// TIA Portal project "Project1" (V20)

(* hardware
DEVICE "S7-1500/ET200MP station_1"  S7-1500 station
   slot 0: "Rail_0"  Rack  6ES7 590-1***0-0AA0
   slot 1: "PLC_2"  CPU 1515F-2 PN  6ES7 515-2FM01-0AB0  V2.9
      slot 3: "CPU display_1"  6ES7591-1BA00-0AA0
      slot 32768: "PROFINET interface_1"  X1
         slot 32769: "Port_1"  X1 P1
         slot 32770: "Port_2"  X1 P2
      slot 33024: "PROFINET interface_2"  X2
         slot 33025: "Port_1"  X2 P1
      slot 34817: "Virtual CP interface port_1"  Virtual CP interface port  Virtual CP interface port
   slot 2: "DI 16x24VDC BA_1"  DI 16x24VDC BA  6ES7 521-1BH10-0AA0  V1.1
   slot 3: "DQ 16x24VDC/0.5A BA_1"  DQ 16x24VDC/0.5A BA  6ES7 522-1BH10-0AA0  V1.1
DEVICE "HMI_1"  KTP700 Basic PN
   slot 0: "HMI_1"  KTP700 Basic PN  6AV2 123-2GB03-0AX0  17.0.0.0
   slot 1: "HMI_RT_1"  KTP700 Basic PN  6AV2 123-2GB03-0AX0  17.0.0.0
   slot 5: "HMI_1.IE_CP_1"  PROFINET Interface  17.0.0.0
      slot 1: "PROFINET Interface_1"  PROFINET Interface
         slot 1: "Port_1"  Port
*)

// ===== PLC "PLC_2"  CPU 1515F-2 PN =====

VAR_GLOBAL   // PLC tag table "Default tag table"
   "KM_Moteur" AT %Q0.0 : Bool;
   "BP_Marche" AT %M0.0 : Bool;
   "BP_Arret_OK" AT %M0.1 : Bool;
   "Niveau_Cuve" AT %MD20 : Real;
   "Vitesse_Pompe" AT %MD24 : Real;
   "Vanne_Vidange" AT %M0.3 : Bool;
   "Cuve_Pleine" AT %M0.2 : Bool;
   "Demande_Production" AT %MD28 : Real;
   "Debit_Sortie" AT %MD32 : Real;
   "Delta_Niveau_Sortie" AT %MD36 : Real;
   "Niveau_Cuve_Calcule" AT %MD40 : Real;
   "Demande_Production_Limitee" AT %MD44 : Real;
   "Debit_Entree" AT %MD48 : Real;
   "Delta_Niveau_Entree" AT %MD52 : Real;
   "Debit_Vidange" AT %MD56 : Real;
   "Autorisation_Vidange" AT %M0.4 : Bool;
   "Debit_Sortie_Total" AT %MD60 : Real;
   "Niveau_Apres_Entree" AT %MD64 : Real;
   "Debit_Entree_Theorique" AT %MD68 : Real;
   "Vitesse_Pompe_Manuelle" AT %MD72 : Real;
END_VAR

DATA_BLOCK "Main_Safety_RTG1_DB"   // DB1, F_DB
{ S7_Optimized_Access := 'TRUE' }
NAME : FUSI
VERSION : 0.1
// stored: InstanceOfName Main_Safety_RTG1
"Main_Safety_RTG1"
BEGIN
END_DATA_BLOCK

DATA_BLOCK "FB_Regulation_Niveau_DB"   // DB3
{ S7_Optimized_Access := 'TRUE' }
VERSION : 0.1
// stored: InstanceOfName FB_Regulation_Niveau
"FB_Regulation_Niveau"
BEGIN
END_DATA_BLOCK

FUNCTION_BLOCK "Main_Safety_RTG1"   // FB1, F_FBD
{ S7_Optimized_Access := 'TRUE' }
BEGIN
END_FUNCTION_BLOCK

FUNCTION_BLOCK "FB_Regulation_Niveau"   // FB2, LAD
{ S7_Optimized_Access := 'TRUE' }
VERSION : 0.1
   VAR
      Consigne_Niveau : Real := 70.0;
      Mode_Auto : Bool;
      Vitesse_PID : Real;
      PID_Actif : Bool;
      Mode_Manuel : Bool;
      Mode_PID : Int := 3;
      Etat_PID : Int;
   END_VAR
BEGIN

REGION Network 1
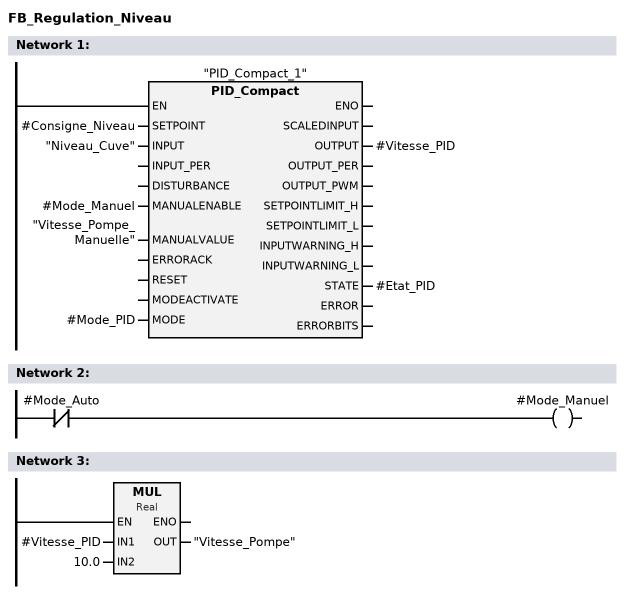
   "PID_Compact_1"(Setpoint := #Consigne_Niveau,   // PID_Compact
                   Input := "Niveau_Cuve",
                   ManualEnable := #Mode_Manuel,
                   ManualValue := "Vitesse_Pompe_Manuelle",
                   Mode := #Mode_PID,
                   Output => #Vitesse_PID,
                   State => #Etat_PID);
END_REGION

REGION Network 2
   RUNG wire#powerrail
      I_Contact( #Mode_Auto )
      Coil( #Mode_Manuel )
   END_RUNG
   // the same network as SCL:
   #Mode_Manuel := NOT #Mode_Auto;
END_REGION

REGION Network 3
   RUNG wire#powerrail
      { S7_Templates := "SrcType := Real" } Mul(in1 := #Vitesse_PID, in2 := 10.0, out => "Vitesse_Pompe")
   END_RUNG
   // the same network as SCL:
   "Vitesse_Pompe" := #Vitesse_PID * 10.0;
END_REGION
END_FUNCTION_BLOCK

ORGANIZATION_BLOCK "Main"   // OB1, LAD, ProgramCycle
TITLE = "Main Program Sweep (Cycle)"
{ S7_Optimized_Access := 'TRUE' }
VERSION : 0.1
   VAR_INPUT
      Initial_Call : Bool;   // Initial call of this OB
      Remanence : Bool;   // =True, if remanent data are available
   END_VAR
BEGIN

REGION Network 1
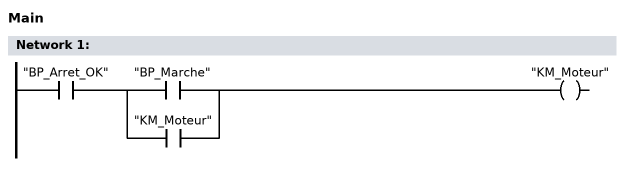
   RUNG wire#powerrail
      Contact( "BP_Arret_OK" )
      wire#w1
      Contact( "BP_Marche" )
      wire#w2
      Coil( "KM_Moteur" )
   END_RUNG
   RUNG wire#w1
      Contact( "KM_Moteur" )
   END_RUNG wire#w2
   // the same network as SCL:
   "KM_Moteur" := "BP_Arret_OK" AND ("BP_Marche" OR "KM_Moteur");
END_REGION
END_ORGANIZATION_BLOCK

ORGANIZATION_BLOCK "OB30_Simulation_Cuve"   // OB30, LAD, CyclicInterrupt
{ S7_Optimized_Access := 'TRUE' }
VERSION : 0.1
   VAR_INPUT
      Initial_Call : Bool;   // Initial call of this OB
      Event_Count : Int;   // Events discarded
   END_VAR
BEGIN

REGION Network 1
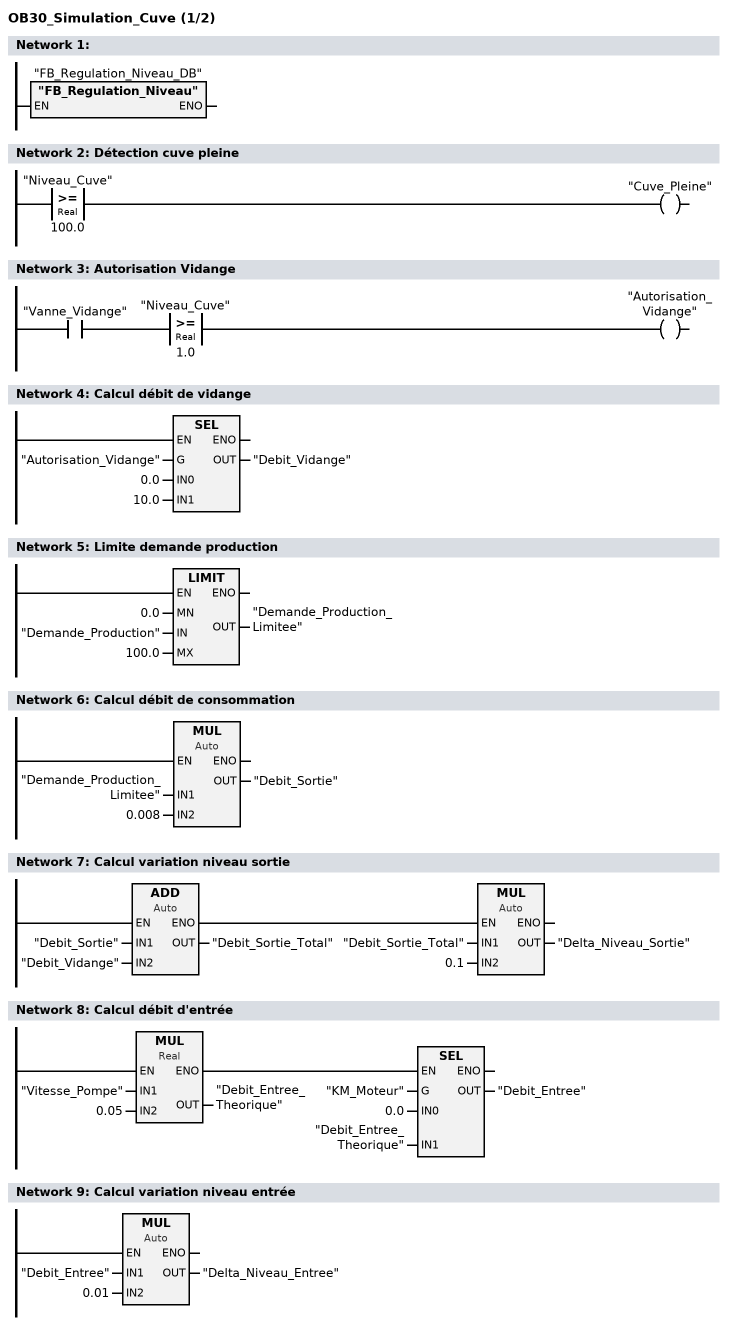
   RUNG wire#powerrail
      "FB_Regulation_Niveau_DB"()
   END_RUNG
   // the same network as SCL:
   "FB_Regulation_Niveau_DB"();   // "FB_Regulation_Niveau"
END_REGION

REGION Network 2: Détection cuve pleine
   RUNG wire#powerrail
      { S7_Templates := "SrcType := Real" } GE_Contact(in1 := "Niveau_Cuve", in2 := 100.0)
      Coil( "Cuve_Pleine" )
   END_RUNG
   // the same network as SCL:
   "Cuve_Pleine" := "Niveau_Cuve" >= 100.0;
END_REGION

REGION Network 3: Autorisation Vidange
   RUNG wire#powerrail
      Contact( "Vanne_Vidange" )
      { S7_Templates := "SrcType := Real" } GE_Contact(in1 := "Niveau_Cuve", in2 := 1.0)
      Coil( "Autorisation_Vidange" )
   END_RUNG
   // the same network as SCL:
   "Autorisation_Vidange" := "Vanne_Vidange" AND ("Niveau_Cuve" >= 1.0);
END_REGION

REGION Network 4: Calcul débit de vidange
   "Debit_Vidange" := SEL(G := "Autorisation_Vidange", IN0 := 0.0, IN1 := 10.0);
END_REGION

REGION Network 5: Limite demande production
   "Demande_Production_Limitee" := LIMIT(MN := 0.0, IN := "Demande_Production", MX := 100.0);
END_REGION

REGION Network 6: Calcul débit de consommation
   RUNG wire#powerrail
      Mul(in1 := "Demande_Production_Limitee", in2 := 0.008, out => "Debit_Sortie")
   END_RUNG
   // the same network as SCL:
   "Debit_Sortie" := "Demande_Production_Limitee" * 0.008;
END_REGION

REGION Network 7: Calcul variation niveau sortie
   RUNG wire#powerrail
      Add(in1 := "Debit_Sortie", in2 := "Debit_Vidange", out => "Debit_Sortie_Total")
      Mul(in1 := "Debit_Sortie_Total", in2 := 0.1, out => "Delta_Niveau_Sortie")
   END_RUNG
   // the same network as SCL:
   "Debit_Sortie_Total" := "Debit_Sortie" + "Debit_Vidange";
   "Delta_Niveau_Sortie" := "Debit_Sortie_Total" * 0.1;
END_REGION

REGION Network 8: Calcul débit d'entrée
   "Debit_Entree_Theorique" := "Vitesse_Pompe" * 0.05;
   "Debit_Entree" := SEL(G := "KM_Moteur", IN0 := 0.0, IN1 := "Debit_Entree_Theorique");
END_REGION

REGION Network 9: Calcul variation niveau entrée
   RUNG wire#powerrail
      Mul(in1 := "Debit_Entree", in2 := 0.01, out => "Delta_Niveau_Entree")
   END_RUNG
   // the same network as SCL:
   "Delta_Niveau_Entree" := "Debit_Entree" * 0.01;
END_REGION

REGION Network 10: Calcul niveau après remplissage
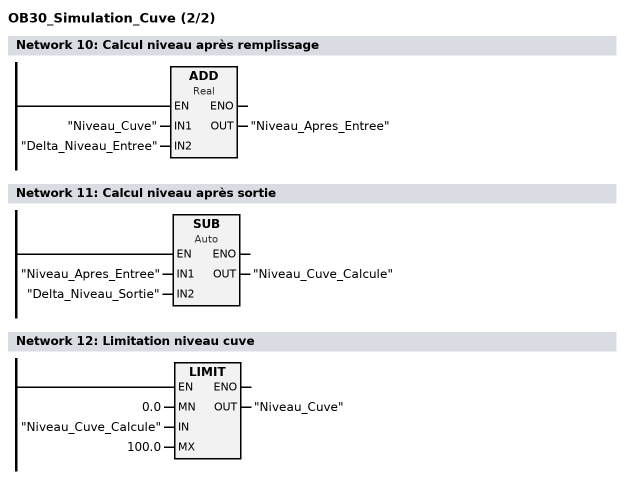
   RUNG wire#powerrail
      { S7_Templates := "SrcType := Real" } Add(in1 := "Niveau_Cuve", in2 := "Delta_Niveau_Entree", out => "Niveau_Apres_Entree")
   END_RUNG
   // the same network as SCL:
   "Niveau_Apres_Entree" := "Niveau_Cuve" + "Delta_Niveau_Entree";
END_REGION

REGION Network 11: Calcul niveau après sortie
   RUNG wire#powerrail
      Sub(in1 := "Niveau_Apres_Entree", in2 := "Delta_Niveau_Sortie", out => "Niveau_Cuve_Calcule")
   END_RUNG
   // the same network as SCL:
   "Niveau_Cuve_Calcule" := "Niveau_Apres_Entree" - "Delta_Niveau_Sortie";
END_REGION

REGION Network 12: Limitation niveau cuve
   "Niveau_Cuve" := LIMIT(MN := 0.0, IN := "Niveau_Cuve_Calcule", MX := 100.0);
END_REGION
END_ORGANIZATION_BLOCK

(* ===== HMI "HMI_RT_1" =====
system functions are stored by id; their names below are inferred from use
connection "HMI_Connection_2": ETHERNET, SMART_S7_1500_OMS
connection "HMI_Connection_3": ETHERNET, SMART_S7_1500_OMS

HMI tags "Default tag table"
   "Vanne_Vidange_HMI" : Bool = PLC Vanne_Vidange AT %M0.3, 1 s
   "BP_Marche" : Bool = PLC BP_Marche AT %M0.0, 1 s
   "BP_Arret_OK" : Bool = PLC BP_Arret_OK AT %M0.1, 1 s
   "KM_Moteur" : Bool = PLC KM_Moteur AT %Q0.0, 1 s
   "Demande_Production_HMI" : Real = PLC Demande_Production AT %MD28, 1 s
   "Niveau_Cuve_HMI" : Real = PLC Niveau_Cuve AT %MD20, 1 s
   "Vitesse_Pompe_Manuelle_HMI" : Real = PLC Vitesse_Pompe_Manuelle AT %MD72, 1 s
   "Mode_Auto_HMI" : Bool = PLC FB_Regulation_Niveau_DB.Mode_Auto AT %DB1.DBX0.0, 1 s
   "Consigne_Niveau_HMI" : Real = PLC FB_Regulation_Niveau_DB.Consigne_Niveau AT %DB1.DBX0.0, 1 s
   "PID_Compact_1_CtrlParamsBackUp_Gain" : Real = PLC PID_Compact_1.CtrlParamsBackUp.Gain, 1 s
   "PID_Compact_1_CtrlParamsBackUp_Ti" : Real = PLC PID_Compact_1.CtrlParamsBackUp.Ti, 1 s
   "PID_Compact_1_Retain_CtrlParams_Gain" : Real = PLC PID_Compact_1.Retain.CtrlParams.Gain, 1 s
   "PID_Compact_1_Retain_CtrlParams_Ti" : Real = PLC PID_Compact_1.Retain.CtrlParams.Ti, 1 s

Template "Template_1" 800x480
   Button "Exit" at 714,429 size 71x50; TextOff 'Exit'; PictureOff "ExitRuntime_KTP700_Basic_DP_TR"; PictureOn "ExitRuntime_KTP700_Basic_DP_TR"
      on Release: StopRuntime(0)
   Button "Template_Button" at 614,429 size 71x50; TextOff 'Text'
   Button "Template_Button_1" at 514,429 size 71x50; TextOff 'Text'
   Button "Template_Button_2" at 414,429 size 71x50; TextOff 'Text'
   Button "Template_Button_3" at 314,429 size 71x50; TextOff 'Text'
   Button "Template_Button_4" at 214,429 size 71x50; TextOff 'Text'
   Button "Alarms" at 114,429 size 71x50; TextOff 'Alarms'; PictureOff "AlarmDisplay_KTP700_Basic_DP_TR"; PictureOn "AlarmDisplay_KTP700_Basic_DP_TR"
      on Release: function_ef3f5d25("Alarm window_Unacknowledged", -1)
   Button "Start screen" at 14,429 size 71x50; TextOff 'Start screen'; PictureOff "NavigateHome_KTP700_Basic_DP_TR"; PictureOn "NavigateHome_KTP700_Basic_DP_TR"
      on Release: ActivateScreen("Root screen", 0)
   SymbolicIOField "Symbolic_IO_Field_Screen" at 93,9 size 600x33; TextOff '0'; TextOn '1'; TextList "TextList_ScreenNames"
      ProcessValue <- "Vanne_Vidange_HMI"
   DateTimeField "HmiScreenItemData" at 695,25 size 105x25
   DateTimeField "HmiScreenItemData_1" at 695,0 size 105x25
   GraphicView "Logo" at 0,0 size 91x51; Picture "Logo of HMI_1"

screen "Root screen" 800x480, template "Template_1"
   on GenerateScreen: SetTag("Vanne_Vidange_HMI", 1)
   TextField "HmiScreenItemData" at 80,225 size 640x25; Text 'Welcome to HMI_1 (KTP700 Basic+ DP)!'

screen "Screen_1" 800x480
   Bar "Bar_1" at 536,85 size 41x217; MinimumValue 0; MaximumValue 100
      ProcessValue <- "Niveau_Cuve_HMI"
   IOField "I/O field_1" at 659,147 size 49x38; FormatPattern 999
      ProcessValue <- "Demande_Production_HMI"
   IOField "I/O field_4" at 85,253 size 96x32; FormatPattern s999999999.999
      ProcessValue <- "Consigne_Niveau_HMI"
   IOField "I/O field_3" at 126,163 size 68x28; FormatPattern s999999999.999
      ProcessValue <- "Vitesse_Pompe_Manuelle_HMI"
   IOField "I/O field_2" at 393,152 size 96x32; FormatPattern s999999999.999
      ProcessValue <- "Niveau_Cuve_HMI"
   Switch "Switch_1" at 126,127 size 57x26; CaptionText 'Switch'; TextOff 'OFF'; TextOn 'ON'
      ProcessValue <- "Mode_Auto_HMI"
   TextField "Text field_2" at 12,127 size 110x20; Text 'AUTO [ON/OFF] :'
   TextField "Text field_3" at 9,163 size 113x20; Text 'MANUAL VALUE :'
   TextField "Text field_4" at 12,253 size 73x20; Text 'SETPOINT :'
   IOField "I/O field_5" at 85,285 size 96x32; FormatPattern s999999999.999
      ProcessValue <- "PID_Compact_1_Retain_CtrlParams_Gain"
   TextField "Text field_5" at 33,291 size 41x20; Text 'Gain :'
   TextField "Text field_6" at 48,317 size 28x20; Text 'Ti :'
   IOField "I/O field_6" at 85,317 size 96x32; FormatPattern s999999999.999
      ProcessValue <- "PID_Compact_1_Retain_CtrlParams_Ti"
   TextField "Text field_7" at 612,93 size 148x23; Text 'WATER DEMAND'
   TextField "Text field_1" at 602,195 size 158x59; Text '0 % No consumption 25 % Low consumption 50 % Medium consumption 75 % High consumption 100 % Maximum consumption'
   TextField "Text field_8" at 39,19 size 164x28; Text 'PUMP SETTINGS'
   TextField "Text field_9" at 55,205 size 128x22; Text 'PI PARAMETERS'
   TextField "Text field_10" at 48,71 size 145x22; Text 'OPERATING MODE'
   Button "Button_1" at 12,436 size 96x32; TextOff 'RUN'
      on Press: SetBit("BP_Marche")
      on Release: ResetBit("BP_Marche")
   Button "Button_2" at 129,437 size 96x32; TextOff 'STOP'
      on Press: ResetBit("BP_Arret_OK")
      on Release: SetBit("BP_Arret_OK")
   Circle "Circle_1" at 76,363 size 67x67
      Appearance <- "KM_Moteur"
   TextField "Text field_11" at 379,399 size 144x23; Text 'DRAIN CONTROL'
   Button "Button_3" at 376,434 size 161x32; TextOff 'OPEN DRAIN'
      on Press: SetBit("Vanne_Vidange_HMI")
      on Release: ResetBit("Vanne_Vidange_HMI")
   TrendView "Trend view_1" at 548,325 size 252x155
*)